TEXTLIST TextList_StateLong
  0 = 'Off'
  1 = 'Standby'
  2 = 'Not Clean'
  3 = 'CIP1 - Rinzed'
  4 = 'CIP2 - Deterged'
  5 = 'CIP3 - Deterged + Clean'
  6 = 'CIP4 - Disinfected'
  7 = 'CIP5 - Done'
  8 = 'Water Ready'
  9 = 'Ready'
  10 = 'Production'
  11 = 'Empty'
  12 = 'Expired'
   = ''
END_TEXTLIST

(* stored: Version 1.1.0.1, ProductVersion 3.1.4024.12
   TextList TextList_StateLong: Id {6452d8ce-591d-49e7-a3a5-3c9025563a85} *)
